ADAPTER mgz (* Adapter Interface *)
  (* Standard: 61499-1 *)
  (* Version 0.0, 10/22/2026, lizar, Schneider Electric *)
  PACKAGE Main;
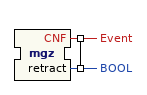
  EVENT_OUTPUT
    CNF WITH retract; (* Confirmation from Plug *)
  END_EVENT
  VAR_OUTPUT
    retract : BOOL; (* Indication Data from Plug *)
  END_VAR
  SERVICE SOCKET/PLUG
    SEQUENCE request_confirm
      SOCKET.REQ(REQD) -> PLUG.REQ(REQD);
      PLUG.CNF(CNFD) -> SOCKET.CNF(CNFD);
    END_SEQUENCE
    SEQUENCE indication_response
      PLUG.IND(retract) -> SOCKET.IND(retract);
      SOCKET.RSP(RSPD) -> PLUG.RSP(RSPD);
    END_SEQUENCE
  END_SERVICE
END_ADAPTER
